# B&R Automation Studio project Lab4
Automation Studio 4.5.2.102; technology packages: Acp10Arnc0 5.2.1

## Configuration Config1

CPU 4PP065.0571-P74, AutomationRuntime D4.52, Build 4.1.2, Vc V4.52.0, Safety 1.6

### Task classes (Cpu.sw)
```
Cyclic#1 (cycle 2000 us, tolerance 0 us):
  ncsdcctrl <- ncsdcctrl.prg
Cyclic#4:
  Program <- Program.prg
DataObjects: Acp10sys
NcDataObjects: acp10etxen <- acp10etxen.dob, gAxis01a <- gAxis01obj.gAxis01a.dob, gAxis01i <- gAxis01obj.gAxis01i.dob
Binaries: udbdef, TCData, vcpfpp30, vcmgr, vcpdpp30, arialbd, vcpdsw, vcalarm, vcshared, vcgclass, Visu01, vctcal, vccbtn, vcfile, vcdsint, Visu03, vcrt, vcpfmtcx, vcbclass, vcfntttf, vcptelo, vcdsloc, vccovl, Visu02, arial, vcctext, vccslider, vcctrend, vccdt, iomap, ashwac, Role, sysconf, arconfig, asfw, User, ashwd, Acp10map, acp10cfg, vccstr, vccbmp
Libraries: Library, Acp10par, NcGlobal, Acp10man, Acp10sdc, Acp10_MC, brsystem, sys_lib, runtime, AsBrStr, fileio, vcresman, dataobj, astime, powerlnk, asieccon
```

### Hardware
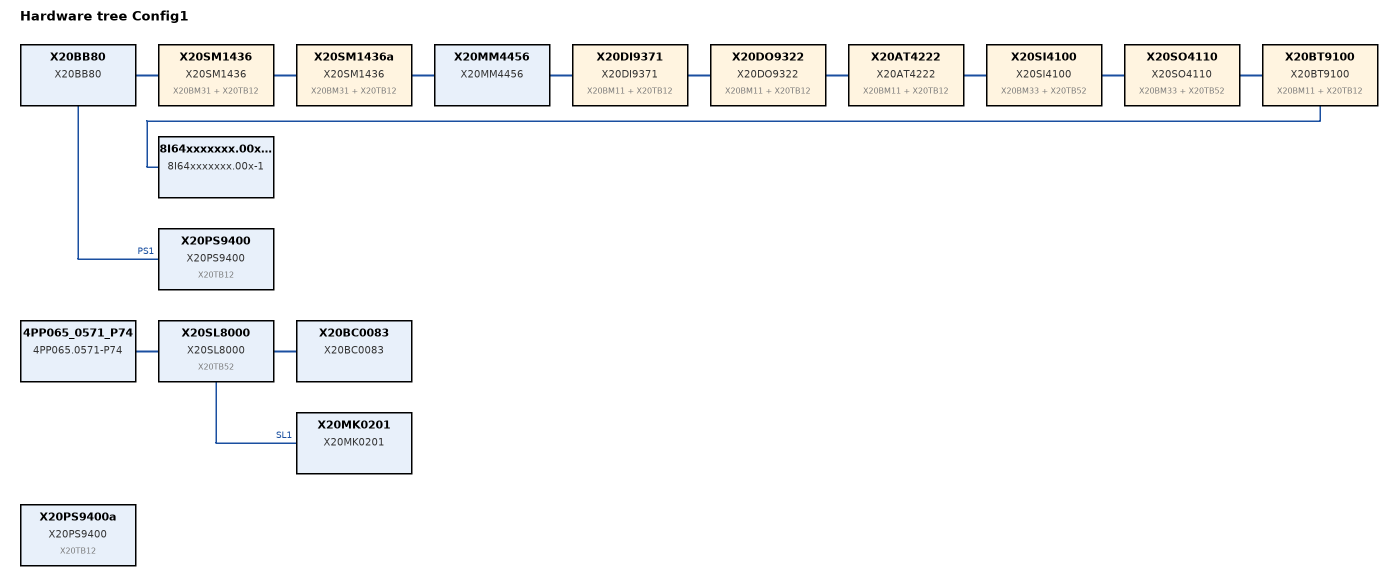
```
4PP065_0571_P74 : 4PP065.0571-P74 v1.1.2.0
  Connector IF4:
    Baudrate = 0
    InaNodeNumber = 1
  Connector IF5:
    ActivateDevice = 1
    Mode = Manual
    InternetAddress = 10.0.1.10
    SubnetMask = 255.255.255.0
    Vnc1
    VncKeyMappingFile1 = VC\PS2-Keyboard.dis
  ConfigurationID = labBR
  TimerDeviceType = EPLX2X
  TimerDevice = 4PP065_0571_P74.IF4
  TaskClassIdleTime = 2000
  Cyclic1Duration = 2000
  Cyclic1Tolerance = 0
  Cyclic1Output = 1
8I64xxxxxxx.00x-1 : 8I64xxxxxxx.00x-1 v2.1.3.0  [X2X1 -> X20BT9100.X2X1 [Cable Type=X2XCable, Length=10, Version=1.0.0.2]]
  packedETAD = packed
  packedCMDD = packed
X20AT4222 : X20AT4222 v1.2.3.0  [SS1 -> X20TB12f.SS; SL -> X20BM11b.SL1]
X20BB80 : X20BB80 v1.0.2.0
X20BC0083 : X20BC0083 v2.9.0.0  [PLK1 -> X20SL8000.PLK2 [Cable Type=PowerlinkCable, Length=10, Version=1.0.0.2]; SL -> X20BB80.SL1]
X20BM11 : X20BM11 v1.0.0.1  [X2X1 -> X20MM4456.X2X2]
X20BM11a : X20BM11 v1.0.0.1  [X2X1 -> X20BM11.X2X2]
X20BM11b : X20BM11 v1.0.0.1  [X2X1 -> X20BM11a.X2X2]
X20BM11c : X20BM11 v1.0.0.1  [X2X1 -> X20BM33a.X2X2]
X20BM31 : X20BM31 v1.0.0.1  [X2X1 -> X20BB80.IF1]
X20BM31a : X20BM31 v1.0.0.1  [X2X1 -> X20BM31.X2X2]
X20BM33 : X20BM33 v1.0.0.4  [X2X1 -> X20BM11b.X2X2]
X20BM33a : X20BM33 v1.0.0.4  [X2X1 -> X20BM33.X2X2]
X20BT9100 : X20BT9100 v1.0.3.0  [SS1 -> X20TB12g.SS; SL -> X20BM11c.SL1]
X20DI9371 : X20DI9371 v1.0.2.0  [SS1 -> X20TB12d.SS; SL -> X20BM11.SL1]
X20DO9322 : X20DO9322 v1.0.3.0  [SS1 -> X20TB12e.SS; SL -> X20BM11a.SL1]
X20MK0201 : X20MK0201 v1.0.0.0  [SL -> X20SL8000.SL1]
X20MM4456 : X20MM4456 v1.1.5.0  [X2X1 -> X20BM31a.X2X2]
X20PS9400 : X20PS9400 v1.8.0.0  [SS1 -> X20TB12.SS; PS -> X20BB80.PS1]
X20PS9400a : X20PS9400 v1.8.0.0  [SS1 -> X20TB12a.SS]
X20SI4100 : X20SI4100 v1.10.1.1  [SS1 -> X20TB52a.SS; SL -> X20BM33.SL1]
X20SL8000 : X20SL8000 v1.6.5.2  [PLK1 -> 4PP065_0571_P74.IF4 [Cable Type=PowerlinkCable, Length=10, Version=1.0.0.2]; PLK2 -> X20BC0083.PLK1 [Cable Type=PowerlinkCable, Length=10, Version=1.0.0.2]; SS1 -> X20TB52.SS]
  SafeProject = SafeLOGIC-1
X20SM1436 : X20SM1436 v2.3.0.0  [SS1 -> X20TB12b.SS; SL -> X20BM31.SL1]
X20SM1436a : X20SM1436 v2.3.0.0  [SS1 -> X20TB12c.SS; SL -> X20BM31a.SL1]
X20SO4110 : X20SO4110 v1.10.1.1  [SS1 -> X20TB52b.SS; SL -> X20BM33a.SL1]
  SafeModuleID = 3
X20TB12 : X20TB12 v1.0.0.0
X20TB12a : X20TB12 v1.0.0.0
X20TB12b : X20TB12 v1.0.0.0
X20TB12c : X20TB12 v1.0.0.0
X20TB12d : X20TB12 v1.0.0.0
X20TB12e : X20TB12 v1.0.0.0
X20TB12f : X20TB12 v1.0.0.0
X20TB12g : X20TB12 v1.0.0.0
X20TB52 : X20TB52 v1.0.0.1
X20TB52a : X20TB52 v1.0.0.1
X20TB52b : X20TB52 v1.0.0.1
```

### IoMap.iom - 4PP065_0571_P74/IoMap.iom
```iecst
VAR_CONFIG
	::Program:EVIRD.STATE AT %IW."8I64xxxxxxx.00x-1".ETAD_Input;
	::Program:EVIRD.COM AT %QW."8I64xxxxxxx.00x-1".CMDD_Output;
	Cyclic#1.gAxis01_DrvIf.iLifeCnt AT %IB."8I64xxxxxxx.00x-1".SDC_LifeCnt;
	Cyclic#1.gAxis01_DrvIf.iDrvOK AT %IX."8I64xxxxxxx.00x-1".ETAD_Input_Bool_02;
	Cyclic#1.gAxis01_DrvIf.oSetTime AT %QW."8I64xxxxxxx.00x-1".SDC_SetTime;
	Cyclic#1.gAxis01_DiDoIf.iLifeCntDriveReady AT %IB."8I64xxxxxxx.00x-1".SDC_LifeCnt;
	Cyclic#1.gAxis01_DiDoIf.iLifeCntDriveEnable AT %IB."8I64xxxxxxx.00x-1".SDC_LifeCnt;
	Cyclic#1.gAxis01_DiDoIf.oDriveEnable AT %QX."8I64xxxxxxx.00x-1".CMDD_Output_Bool_00;
	Cyclic#1.gAxis01_ModuleOk AT %QX."8I64xxxxxxx.00x-1".CMDD_Output_Bool_01;
	Cyclic#1.gAxis01_ModuleOk AT %QX."8I64xxxxxxx.00x-1".CMDD_Output_Bool_02;
	Cyclic#1.gAxis01_ModuleOk AT %IX."8I64xxxxxxx.00x-1".ModuleOk;
	Cyclic#1.gAxis01_DiDoIf.oDriveEnable AT %QX."8I64xxxxxxx.00x-1".CMDD_Output_Bool_03;
	Cyclic#1.gAxis01_DiDoIf.iDriveReady AT %IX."8I64xxxxxxx.00x-1".ETAD_Input_Bool_02;
	::Program:LedState.led1 AT %QX."X20DO9322".DigitalOutput02;
	::Program:LedState.led2 AT %QX."X20DO9322".DigitalOutput03;
	::Program:LedState.led3 AT %QX."X20DO9322".DigitalOutput04;
	::Program:LedState.led4 AT %QX."X20DO9322".DigitalOutput05;
	::Program:DoorState.sw1 AT %IX."X20DI9371".DigitalInput02;
	::Program:DoorState.sw2 AT %IX."X20DI9371".DigitalInput03;
	::Program:DoorState.sw3 AT %IX."X20DI9371".DigitalInput04;
	::Program:DoorState.sw4 AT %IX."X20DI9371".DigitalInput05;
	::Program:DoorState.direction AT %IX."X20DI9371".DigitalInput01;
	 ::Program:DoorState.speed AT %QW."8I64xxxxxxx.00x-1".LFRD_Output;
END_VAR
```

### Acp10cfg.ncc - 4PP065_0571_P74/Motion/Acp10cfg.ncc
```
NcConfiguration (Version=5.02.1, NcSwId=Acp10)
  ACP10CF1_typ:
    cnt_nettrc_rec_drive = 150
    bufsize_trace_upload = 1200
    tc_nc_man_task = Cyclic #1
    glob_pv_as_ncobject = Yes
    ncsys_dl_broadcast = Yes
    ncsys_dl_acp_reset = Yes
    safemc_log_err_to_ax = Yes
    network_init:
      ncsw_init_execute = Yes
      automatic_execute = No
      node_nr_warning = Yes
      net_err_before_ncact = Yes
    nettrc:
      enter_parsecrec = Yes
      enter_ncaction = Yes
      save_ring_startidx = No
    cam_prof_download:
      cam_dat_dl_parallel = No
      tc_cam_dl_parallel = Task class for NC Manager task
    sdc_if[0]:
      if_name = SDC_IF1
      mc_broadcast_size = 800
      mc_broadcast_extdat = No
```

### Acp10map.ncm - 4PP065_0571_P74/Motion/Acp10map.ncm
```
NcMapping (NcSwId=Acp10)
  NcObject gAxis01 (ModuleId=8I64xxxxxxx.00x-1, ModuleAddress=SDC_IF1.ST1, Type=ncAXIS, Channel=1, AcoposSimulation=Off, InitParameter=gAxis01i, AcoposParameter=gAxis01a, Disabled=FALSE, ModuleDisabled=FALSE)
```

## Logical view

Binary libraries used (declarations not repeated): operator, runtime, astime, AsIecCon, Acp10par 5.02.1, NcGlobal 5.02.1, Acp10man 5.02.1, Acp10sdc 5.02.1, Acp10_MC 5.02.1, brsystem, sys_lib, AsBrStr

### Global.var - Global variables
```iecst
VAR
	direction : BOOL := FALSE;
	gAxis01 : ACP10AXIS_typ;
	gAxis01_DiDoIf : SdcDiDoIf_typ := (0);
	gAxis01_DrvIf : SdcDrvIf16_typ := (0);
	gAxis01_HW : SdcHwCfg_typ := (0);
	gAxis01_ModuleOk : BOOL := 0;
	speed : INT;
END_VAR
```

### Package Logical/Libraries - Global libraries

### Library Logical/Libraries/Library (ANSIC)

#### Library.fun
```iecst
{REDUND_ERROR} FUNCTION_BLOCK DriveStateMachine (*TODO: Add your comment here*) (*$GROUP=User,$CAT=User,$GROUPICON=User.png,$CATICON=User.png*)
	VAR_INPUT
		ENABLE : BOOL;
		STATE : UINT;
	END_VAR
	VAR_OUTPUT
		COM : UINT;
	END_VAR
END_FUNCTION_BLOCK

{REDUND_ERROR} FUNCTION_BLOCK DoorStateMachine (*TODO: Add your comment here*) (*$GROUP=User,$CAT=User,$GROUPICON=User.png,$CATICON=User.png*)
	VAR
		swp1 : BOOL := 0;
		swp2 : BOOL := 0;
		swp3 : BOOL := 0;
	END_VAR
	VAR_INPUT
		swp4 : {REDUND_UNREPLICABLE} BOOL := 0;
		sw1 : {REDUND_UNREPLICABLE} BOOL;
		sw2 : {REDUND_UNREPLICABLE} BOOL;
		sw3 : {REDUND_UNREPLICABLE} BOOL;
		sw4 : {REDUND_UNREPLICABLE} BOOL;
		direction : {REDUND_UNREPLICABLE} BOOL;
		state : INT := 0;
	END_VAR
	VAR_OUTPUT
		speed : {REDUND_UNREPLICABLE} INT;
		state_out : INT;
	END_VAR
END_FUNCTION_BLOCK

{REDUND_ERROR} FUNCTION_BLOCK LedStateMachine (*TODO: Add your comment here*) (*$GROUP=User,$CAT=User,$GROUPICON=User.png,$CATICON=User.png*)
	VAR_INPUT
		state : {REDUND_UNREPLICABLE} INT := 0;
	END_VAR
	VAR_OUTPUT
		led1 : {REDUND_UNREPLICABLE} BOOL;
		led2 : {REDUND_UNREPLICABLE} BOOL;
		led3 : {REDUND_UNREPLICABLE} BOOL;
		led4 : {REDUND_UNREPLICABLE} BOOL;
	END_VAR
	VAR
		timer : UINT;
	END_VAR
END_FUNCTION_BLOCK
```

#### DriveStateMachine.c
```c
#include <bur/plctypes.h>
#ifdef __cplusplus
	extern "C"
	{
#endif
	#include "Library.h"
#ifdef __cplusplus
	};
#endif
/* TODO: Add your comment here */
void DriveStateMachine(struct DriveStateMachine* inst)
{
	UINT mask=inst->STATE & 0x6f;
	if (!inst->ENABLE)
	{
		inst->COM = CMD_SHUTDOWN;
	}
	else
	{

		switch (mask)
		{
			case STATE_DISABLED:
				inst->COM=CMD_SHUTDOWN;
				break;

			case STATE_READY:
       			inst->COM=CMD_ENABLED;
				break;

			case STATE_SWITCHED_ON:
       			inst->COM=CMD_SWITCHED_ON;
				break;
		}

	}

	/*TODO: Add your code here*/
}
```

#### DoorStateMachine.c
```c
#include <bur/plctypes.h>
#ifdef __cplusplus
	extern "C"
	{
#endif
#include "Library.h"
#ifdef __cplusplus
	};
#endif
/* State mashine for door control */
void DoorStateMachine(struct DoorStateMachine* inst)
{
	int high = 250;
	int mid = 750;
	int low = 250;
	int false = 0;
	int true = 1;
	switch(inst->state)
	{
		case 0:
			{
				inst->state = 1;
				break;
			}
		case 1:
			if (inst->direction==false && inst->sw1!=inst->swp1){
				inst->state = 2;
				inst->speed = 0;
				break;
			}
			if (inst->direction==true && inst->sw4!=inst->swp4){
				inst->state = 3;
				inst->speed = 0;
				break;
			}
			break;
		case 2:
			if (inst->direction==false){
				inst->state = 4;
				inst->speed = low;
				break;
			}
			break;
		case 3:
			if (inst->direction==true){
				inst->state = 5;
				inst->speed = -low;
				break;
			}
			break;
		case 4:
			if (inst->sw2!=inst->swp2){
				inst->state = 6;
				inst->speed = mid;
				break;
			}
			if (inst->direction==true){
				inst->state = 9;
				inst->speed = -high;
				break;
			}
			break;
		case 5:
			if (inst->sw3!=inst->swp3){
				inst->state = 7;
				inst->speed = -mid;
				break;
			}
			if (inst->direction==false){
				inst->state = 8;
				inst->speed = high;
				break;
			}
			break;
		case 6:
			if (inst->sw3!=inst->swp3){
				inst->state = 8;
				inst->speed = high;
				break;
			}
			if (inst->direction==true){
				inst->state = 7;
				inst->speed = -mid;
				break;
			}
			break;
		case 7:
			if (inst->sw2!=inst->swp2){
				inst->state = 9;
				inst->speed = -high;
				break;
			}
			if (inst->direction==false){
				inst->state = 6;
				inst->speed = mid;
				break;
			}
			break;
		case 8:
			if (inst->sw4!=inst->swp4){
				inst->state = 3;
				inst->speed = 0;
				break;
			}
				break;
		case 9:
			if (inst->sw1!=inst->swp1){
				inst->state = 2;
				inst->speed = 0;
				break;
			}

	}
	inst->state_out = inst->state;
	inst->swp1 = inst->sw1;
	inst->swp2 = inst->sw2;
	inst->swp3 = inst->sw3;
	inst->swp4 = inst->sw4;
	/*TODO: Add your code here*/
}
```

#### LedStateMachine.c
```c
#include <bur/plctypes.h>
#ifdef __cplusplus
	extern "C"
	{
#endif
#include "Library.h"
#ifdef __cplusplus
	};
#endif
/* Tut mog bit vash commentariy */
void LedStateMachine(struct LedStateMachine* inst)
{

	switch(inst->state){
		case 0:
			inst->led1 = 0;
			inst->led1 = 0;
			inst->led1 = 0;
			inst->led1 = 0;
			break;
		case 1:
			if (inst->timer < 5){
				inst->led1 = 0;
				inst->led2 = 0;
				inst->led3 = 0;
				inst->led4 = 0;
				inst->timer = inst->timer + 1;
				break;
			}
			if (inst->timer < 10){
				inst->led1 = 1;
				inst->led2 = 1;
				inst->led3 = 1;
				inst->led4 = 1;
				inst->timer = inst->timer + 1;
				break;
			}
			inst->timer = 0;
			break;
		case 2:
			inst->led1 = 0;
			inst->led2 = 0;
			inst->led3 = 0;
			inst->led4 = 0;
			break;
		case 3:
			inst->led1 = 1;
			inst->led2 = 1;
			inst->led3 = 1;
			inst->led4 = 1;
			break;
		case 4:
			inst->led1 = 1;
			inst->led2 = 0;
			inst->led3 = 0;
			inst->led4 = 0;
			break;
		case 5:
			inst->led1 = 1;
			inst->led2 = 1;
			inst->led3 = 1;
			inst->led4 = 0;
			break;

		case 6:
			inst->led1 = 1;
			inst->led2 = 1;
			inst->led3 = 0;
			inst->led4 = 0;
			break;
		case 7:
			inst->led1 = 1;
			inst->led2 = 1;
			inst->led3 = 0;
			inst->led4 = 0;
			break;
		case 8:
			inst->led1 = 1;
			inst->led2 = 1;
			inst->led3 = 1;
			inst->led4 = 0;
			break;
		case 9:
			inst->led1 = 1;
			inst->led2 = 0;
			inst->led3 = 0;
			inst->led4 = 0;
			break;

	}
}
```

#### Constant.var
```iecst
VAR CONSTANT
	CMD_SWITCHED_ON : UINT := 7;
	CMD_DISABLE_VOLTAGE : UINT := 0;
	CMD_ENABLED : UINT := 15;
	CMD_SHUTDOWN : UINT := 6;
	STATE_READY : UINT := 33;
	STATE_DISABLED : UINT := 64;
	STATE_SWITCHED_ON : UINT := 35;
END_VAR
```

### Program Logical/Program (ANSIC)

#### Main.c - Init, cyclic, exit code
```c
#include <bur/plctypes.h>

#ifdef _DEFAULT_INCLUDES
	#include <AsDefault.h>
	#include <stdlib.h>

#endif

void _INIT ProgramInit(void)
{
	EVIRD.ENABLE = 1;
	LedState.state = DoorState.state_out;

}

void _CYCLIC ProgramCyclic(void)
{
	DriveStateMachine(&EVIRD);
	DoorStateMachine(&DoorState);
	LedState.state = DoorState.state_out;
	LedStateMachine(&LedState);

}

void _EXIT ProgramExit(void)
{

}
```

#### Variables.var - Local variables
```iecst
VAR
	DoorState : DoorStateMachine;
	EVIRD : DriveStateMachine;
	LedState : LedStateMachine;
END_VAR
```

### Program Logical/Gogram (ANSIC)

#### Main.c - Init, cyclic, exit code
```c
#include <bur/plctypes.h>

#ifdef _DEFAULT_INCLUDES
#include <AsDefault.h>
#endif

void _INIT ProgramInit(void)
{
	led_1 = 1;
	led_2 = 0;
	k = 0;
}

void _CYCLIC ProgramCyclic(void)
{
	if(k <4)
	{
		led_1 = !led_1;

	}
	k++;
	if (k ==7)
	{
		k = 0;
	}
	led_2 = !led_2;
}

void _EXIT ProgramExit(void)
{

}
```

#### Variables.var - Local variables
```iecst
VAR
	k : USINT;
END_VAR
```

### Program Logical/ncsdcctrl (IEC)

#### ncsdcctrlCyclic.st
```iecst
PROGRAM _CYCLIC

(* ### BEGIN gAxis01 ### *)

(* life counter emulation of digital inputs *)
        gAxis01_DiDoIf.iLifeCntReference := gAxis01_DiDoIf.iLifeCntReference + 1;
        gAxis01_DiDoIf.iLifeCntNegHwEnd  := gAxis01_DiDoIf.iLifeCntNegHwEnd  + 1;
        gAxis01_DiDoIf.iLifeCntPosHwEnd  := gAxis01_DiDoIf.iLifeCntPosHwEnd  + 1;

(* ### END gAxis01 ### *)

END_PROGRAM
```

#### ncsdcctrlInit.st
```iecst
PROGRAM _INIT

(* ### BEGIN gAxis01 ### *)

(* initialize variables *)
        gAxis01_HW.DrvIf_Typ := ncSDC_DRVSERVO16;
        brsstrcpy(ADR(gAxis01_HW.DrvIf_Name[0]), ADR('gAxis01_DrvIf'));
        gAxis01_HW.DiDoIf_Typ := ncSDC_DIDO;
        brsstrcpy(ADR(gAxis01_HW.DiDoIf_Name[0]), ADR('gAxis01_DiDoIf'));

(* force variable offset generation *)
        gAxis01.size                      := gAxis01.size;
        gAxis01_DrvIf.iLifeCnt            := gAxis01_DrvIf.iLifeCnt;
        gAxis01_DiDoIf.iLifeCntDriveReady := gAxis01_DiDoIf.iLifeCntDriveReady;
        gAxis01_ModuleOk                  := gAxis01_ModuleOk;

(* assign your hardware inputs here*)

(*      gAxis01_DiDoIf.iPosHwEnd  := gAxis01_DiDoIf.iPosHwEnd;
        gAxis01_DiDoIf.iNegHwEnd  := gAxis01_DiDoIf.iNegHwEnd;
        gAxis01_DiDoIf.iReference := gAxis01_DiDoIf.iReference;
 *)

(* ### END gAxis01 ### *)

END_PROGRAM
```

### Data object Logical/acp10etxen (Ett)

- acp10etxen.ett (not shown)

### Package Logical/gAxis01obj - gAxis01obj

### Data object Logical/gAxis01obj/gAxis01a (Apt)

#### gAxis01a.apt
```
AcoposParameterTable:
  Root Parameters:
    230 = PCTRL_S_SET (Name=PCTRL_S_ACT_PARID)
    64201 = 546116.666666667 (Name=SERVO_V_MAX_OUTPUT)
```

### Data object Logical/gAxis01obj/gAxis01i (Ax)

#### gAxis01i.ax
```
InitParameter (Version=5.2.1, NcSwId=Acp10)
  ACP10AXIS_typ:
    dig_in:
      level:
        reference = ncACTIV_HI
        pos_hw_end = ncACTIV_LO
        neg_hw_end = ncACTIV_LO
        trigger1 = ncACTIV_HI
        trigger2 = ncACTIV_LO + ncQUICKSTOP
    encoder_if:
      parameter:
        count_dir = ncSTANDARD
        scaling:
          load:
            units = 1000
            rev_motor = 1
    limit:
      parameter:
        v_pos = 10000
        v_neg = 10000
        a1_pos = 50000
        a2_pos = 50000
        a1_neg = 50000
        a2_neg = 50000
        t_jolt = 0
        t_in_pos = 0
        pos_sw_end = 2000000000
        neg_sw_end = -2000000000
        ds_warning = 500
        ds_stop = 1000
        a_stop = 1.0e30
        dv_stop = 0
        dv_stop_mode = ncOFF
    controller:
      mode = ncPOSITION
      position:
        kv = 50
        tn = 0
        t_predict = 0.01
        t_total = 0.01
        p_max = 1.0e30
        i_max = 0
      speed:
        kv = 2.0
        tn = 0
        t_filter = 0.0
        isq_filter1:
          type = ncOFF
          a0 = 0.0
          a1 = 0.0
          b0 = 0.0
          b1 = 0.0
          b2 = 0.0
          c0_par_id = 0
          c1_par_id = 0
        isq_filter2:
          type = ncOFF
          a0 = 0.0
          a1 = 0.0
          b0 = 0.0
          b1 = 0.0
          b2 = 0.0
          c0_par_id = 0
          c1_par_id = 0
        isq_filter3:
          type = ncOFF
          a0 = 0.0
          a1 = 0.0
          b0 = 0.0
          b1 = 0.0
          b2 = 0.0
          c0_par_id = 0
          c1_par_id = 0
      uf:
        type = ncLINEAR + ncCORRECTION
        auto_config = ncMOTOR_PAR
        u0 = 0
        un = 0
        fn = 50.0
        k_f_slip = 0
      ff:
        torque_load = 0.0
        torque_pos = 0.0
        torque_neg = 0.0
        kv_torque = 0.0
        inertia = 0.0
        t_filter_a = 0.0
    move:
      stop:
        parameter[0]:
          decel_ramp = ncA_LIMIT
          controller = ncON
        parameter[1]:
          decel_ramp = ncA_LIMIT
          controller = ncON
        parameter[2]:
          decel_ramp = ncA_LIMIT
          controller = ncON
        parameter[3]:
          decel_ramp = ncA_LIMIT
          controller = ncON
        quickstop:
          decel_ramp = ncA_LIMIT
          t_jolt = 0
        drive_error:
          decel_ramp = ncA_LIMIT
      homing:
        parameter:
          s = 0
          v_switch = 5000
          v_trigger = 500
          a = 50000
          mode = ncDIRECT
          edge_sw = ncPOSITIVE
          start_dir = ncPOSITIVE
          trigg_dir = ncPOSITIVE
          ref_pulse = ncOFF
          fix_dir = ncOFF
          tr_s_block = 0
          torque_lim = 0
          ds_block = 0
          ds_stop = 0
      basis:
        parameter:
          v_pos = 5000
          v_neg = 5000
          a1_pos = 50000
          a2_pos = 50000
          a1_neg = 50000
          a2_neg = 50000
    message:
      text:
        parameter:
          format = ncBREAK
          columns = 80
          data_modul = acp10etxen
```
